// TRUE while the shared Az/El brake must be commanded closed (MONETcommon#121): the elevation axis is disabled.
// With the elevation disabled and the brake open nothing holds the telescope, which swings if it is unbalanced.
// The brake close in HalfBROT FB_ElevationControl is edge-only (falling edge of bEnable) and bOpenBrake of the
// hydraulics is a latch, so a brake that opens later (manual-mode latch, ADS write, pendant) stayed open.
// Only called in automatic: in manual the azimuth needs the brake open with the elevation disabled.
// Exception (#151): in the Wake&Shake window the drives run their own command with the brake released and the axes not
// enabled by the PLC, so the brake that the operator opened is left open (F_WakeShakeWindow bounds the window).
// #155: the operator may also open it in the window with an elevation error latched. Four level blocks close it while
// they hold (they do not end the window): E-stop, hydraulics error, safety error, covers not open.
FUNCTION F_BrakeMustClose : BOOL
VAR_INPUT
	bElevationEnabled	: BOOL;		// fbElevation.bEnable
	bWakeShakeWindow	: BOOL;		// F_WakeShakeWindow
	bEstop				: BOOL;		// bEstopTriggered
	bHydraulicsError	: BOOL;		// fbHydraulics.Error
	bSafetyError		: BOOL;		// bSafetyError (SafetyHandling.error)
	bCoversOpen			: BOOL;		// fbCovers.Opened
END_VAR

F_BrakeMustClose := NOT bElevationEnabled AND
	(NOT bWakeShakeWindow OR bEstop OR bHydraulicsError OR bSafetyError OR NOT bCoversOpen);

END_FUNCTION

(* stored: Version 1.1.0.1, ProductVersion 3.1.4024.15
   POU F_BrakeMustClose: Id {c15d8543-9f0c-4859-861e-c979b4be4202}, SpecialFunc None *)
